FUNCTION_BLOCK ABSTRACT TestBase
VAR
    _CheckCount  : INT;
    _FailedCount : INT;
    _LastFailure : STRING(255);
END_VAR
(*
    TestBase

    Shared bookkeeping for framework-free tests. A derived test implements
    Run() and calls Check() for everything it wants to verify.
*)

METHOD PUBLIC ABSTRACT Run
END_METHOD

METHOD PROTECTED Check
VAR_INPUT
    Condition : BOOL;
    Message   : STRING(255);    // what should be true, not what went wrong
END_VAR
_CheckCount := _CheckCount + 1;
IF NOT Condition THEN
    _FailedCount := _FailedCount + 1;
    _LastFailure := Message;
END_IF
END_METHOD

PROPERTY PUBLIC HasPassed : BOOL
GET
HasPassed := _CheckCount > 0 AND _FailedCount = 0;
END_GET
END_PROPERTY

PROPERTY PUBLIC FailedCount : INT
GET
FailedCount := _FailedCount;
END_GET
END_PROPERTY

PROPERTY PUBLIC LastFailure : STRING(255)
GET
LastFailure := _LastFailure;
END_GET
END_PROPERTY

END_FUNCTION_BLOCK

(* stored: Version 1.1.0.1, ProductVersion 3.1.4026.0
   POU TestBase: Id {00d9475d-5935-4b0d-a71b-28a102aa94b4}, SpecialFunc None
   Method Run: Id {4c16e47f-57f9-412a-8ad0-d28ec9a619a6}
   Method Check: Id {c6242960-d1b8-4a18-be43-d329ebe3b52b}
   Property HasPassed: Id {4e595662-ae47-4cfc-8a1c-27a0ca77691a}
   Get Get: Id {fa494ea5-fe5b-44dd-ad83-4cc0bad07c3f}
   Property FailedCount: Id {787a173b-d7bd-4af3-a47a-03a7371f1103}
   Get Get: Id {2e6372e1-7eba-4f14-9c6c-b7cf27dfbd5a}
   Property LastFailure: Id {0ae27779-fd5b-4f61-b1d2-44d4cb5fcf95}
   Get Get: Id {254a139e-d29a-4440-812a-ca0016b9e6d3} *)
